INTERFACE iSwitch

PROPERTY PUBLIC IsPressed : BOOL
GET
END_GET
END_PROPERTY

PROPERTY IsReleased : BOOL
GET
END_GET
END_PROPERTY

END_INTERFACE

(* stored: Version 1.1.0.1
   Itf iSwitch: Id {2b8cdf8a-a619-4e44-ba18-5ff28feae6d7}
   Property IsPressed: Id {76e8bbdf-c484-4aa9-82c0-6b7f3dc3327a}
   Get Get: Id {b1befc1a-e193-4b1a-b19b-81d2f9e2197e}
   Property IsReleased: Id {72547f3f-78f0-4e28-87f6-c436549bb588}
   Get Get: Id {b83f7f50-cdcf-4a72-8eba-03891819d814} *)
